Fanuc KAREL source: kd00074.KL

-- PROVISIONAL review KL for V770-1; original PC SHA256 bfcb592e1e3c5de7c206587bf5d3ec796506749b2604cc6cb08b347ca98317c8
-- Incomplete behavior may be omitted. Consult companion uncertainty JSON. Do not deploy.
PROGRAM KD00074
%NOLOCKGROUP
VAR
  I : INTEGER
  J : INTEGER
  B : BOOLEAN
  R : REAL
  S : STRING[80]
BEGIN
  -- UNRESOLVED_PC offsets 5-7; opcodes 9C,3B
  -- UNRESOLVED_PC offsets 12-16; opcodes 7F
END KD00074
